Fanuc KAREL source: kc00001.KL

-- PROVISIONAL review KL for V770-1; original PC SHA256 c0c4265d8e1ea12dd41e54b34e7da74230b03fe169aaa3a1394c3efa7db0a061
-- Incomplete behavior may be omitted. Consult companion uncertainty JSON. Do not deploy.
PROGRAM KC00001
%NOLOCKGROUP
BEGIN
  -- UNRESOLVED_PC offsets 5-14; opcodes 3F,75
  -- UNRESOLVED_PC offsets 19-28; opcodes 3F,75
  -- UNRESOLVED_PC offsets 33-71; opcodes 27,22,22,22,2A,22,2A,22,31
  -- UNRESOLVED_PC offsets 76-80; opcodes 7F
END KC00001
